(* IEC 61131-3 sources: trust-platform/examples/communication/ads_line1/src, 2 files *)

(* ---- config.st ---- *)
CONFIGURATION Config
RESOURCE CommRes ON PLC
    TASK MainTask (INTERVAL := T#100ms, PRIORITY := 1);
    PROGRAM Main WITH MainTask : Main;
END_RESOURCE
END_CONFIGURATION

(* ---- main.st ---- *)
PROGRAM Main
VAR_EXTERNAL
    line1_temp : REAL;
    line1_ready : BOOL;
    line1_setpoint : REAL;
    line1_status : WORD;
    line1_temp_quality : ADS_QUALITY;
END_VAR

IF line1_ready THEN
    line1_setpoint := line1_temp;
ELSE
    line1_setpoint := REAL#0.0;
END_IF;
END_PROGRAM
